TYPE (* Identification of a module on a modular EtherCAT slave *)
  (* Description: Copyright (c) 2026 Sichuan Qunyuan Technology Co., Ltd. This program and the accompanying materials are made available under the terms of the Eclipse Public License 2.0 which is available at https://www.eclipse.org/legal/epl-2.0/ SPDX-License-Identifier: EPL-2.0 *)
  (* Version 1.0, 2026-04-14, Zijun Tang *)
  PACKAGE eclipse4diac::io::ethercat;
  ECModuleConfig : STRUCT
    ModuleIdent : UDINT; (* ESI Modules/Module Type/@ModuleIdent *)
    Slot : UINT; (* Slot index on the modular device *)
  END_STRUCT;
END_TYPE
